FUNCTION_BLOCK logiBUS_QDA_FREQ (* Composite FB for a frequency output (MCPWM, duty cycle 50 %, frequency in mHz in DWORD) *)
  (* Standard: 61499-2; Description: Copyright (c) 2026 HR Agrartechnik GmbH This program and the accompanying materials are made available under the terms of the Eclipse Public License 2.0 which is available at https://www.eclipse.org/legal/epl-2.0/ SPDX-License-Identifier: EPL-2.0 *)
  (* Version 1.0, 2026-11-06, Franz Höpfinger, HR Agrartechnik GmbH, initial version *)
  PACKAGE logiBUS::io::DQ;
  IMPORT logiBUS::io::DQ::logiBUS_DO::Invalid;
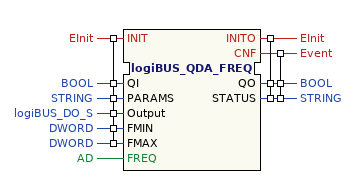
  EVENT_INPUT
    INIT : EInit WITH QI, PARAMS, Output, FMIN, FMAX; (* Service Initialization *)
  END_EVENT
  EVENT_OUTPUT
    INITO : EInit WITH QO, STATUS; (* Initialization Confirm *)
    CNF WITH QO, STATUS; (* Confirmation of Requested Service *)
  END_EVENT
  VAR_INPUT
    QI : BOOL; (* Event Input Qualifier *)
    PARAMS : STRING; (* Service Parameters *)
    Output : logiBUS::io::DQ::logiBUS_DO_S := Invalid; (* Identify the Output Output_Q1..Q8 *)
    FMIN : DWORD := 10000; (* Lowest frequency in mHz, read at INIT. Sets the timer resolution (16-bit timer: resolution = about FMIN * 65536): the higher FREQ is above FMIN, the coarser the steps (step about FREQ^2 / resolution). Default 10 Hz: 640 kHz resolution, step 1.6 Hz at 1 kHz, 156 Hz at 10 kHz *)
    FMAX : DWORD := 10000000; (* Highest frequency in mHz, read at INIT. FREQ above it is limited. Never more than the chip can produce with the resolution from FMIN (half the resolution) *)
  END_VAR
  VAR_OUTPUT
    QO : BOOL; (* Event Output Qualifier *)
    STATUS : STRING; (* Service Status *)
  END_VAR
  SOCKETS
    FREQ : adapter::types::unidirectional::AD; (* Frequency in mHz (D1, 1000 = 1 Hz, 0 = off) like ISOBUS DDI 583 *)
  END_SOCKETS
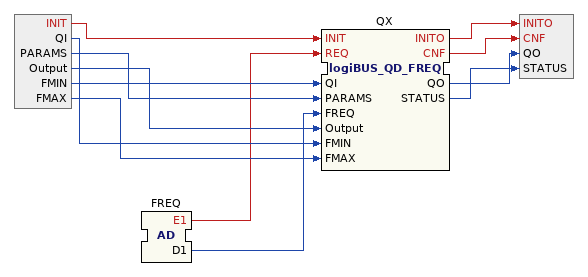
  FBS
    QX : logiBUS::io::DQ::logiBUS_QD_FREQ;
  END_FBS
  EVENT_CONNECTIONS
    INIT TO QX.INIT;
    QX.INITO TO INITO;
    FREQ.E1 TO QX.REQ;
    QX.CNF TO CNF;
  END_CONNECTIONS
  DATA_CONNECTIONS
    FREQ.D1 TO QX.FREQ;
    QI TO QX.QI;
    PARAMS TO QX.PARAMS;
    QX.QO TO QO;
    QX.STATUS TO STATUS;
    Output TO QX.Output;
    FMIN TO QX.FMIN;
    FMAX TO QX.FMAX;
  END_CONNECTIONS
END_FUNCTION_BLOCK
